FUNCTION_BLOCK LimiterTemp (* Basic Function Block Type *)
  (* Standard: 61499-2 *)
  (* Version 0.0, 6/22/2016, Andrei, nxtControl GmbH, Template *)
  PACKAGE Main;
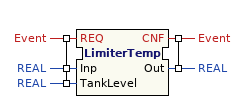
  EVENT_INPUT
    REQ WITH Inp, TankLevel; (* Normal Execution Request *)
  END_EVENT
  EVENT_OUTPUT
    CNF WITH Out; (* Execution Confirmation *)
  END_EVENT
  VAR_INPUT
    Inp : REAL; (* Input event qualifier *)
    TankLevel : REAL;
  END_VAR
  VAR_OUTPUT
    Out : REAL; (* Output event qualifier *)
  END_VAR
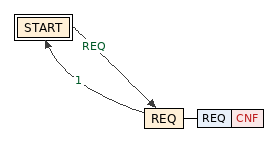
  EC_STATES
    START; (* Initial State *)
    REQ : REQ -> CNF; (* Normal execution *)
  END_STATES
  EC_TRANSITIONS
    START TO REQ := REQ;
    REQ TO START := 1;
  END_TRANSITIONS
  ALGORITHM REQ IN ST: (* Normally executed algorithm *)
IF (Inp > 100.0) AND (TankLevel>1.0) THEN
	Out := 100.0;
ELSIF (Inp <= 100.0) AND (TankLevel>1.0) THEN
	Out := Inp;
ELSE
	Out := 20.0;
END_IF;
  END_ALGORITHM
END_FUNCTION_BLOCK
